(* IEC 61131-3 sources: guidance-for-physical-ai-production-designer-on-aws/source/plan2cell/crates/bt2plc/tests/golden/welding_cell_2_small/codesys/head/GVL, 2 files *)

(* ---- GVL_Cell.st ---- *)
(*
 * GVL_Cell - generated by bt2plc 0.1.0 - DO NOT EDIT
 * Plan   : bt_1790934549_welding_cell_2_small (cell welding_cell_2_small)
 * Grants : planned ticket order
 * IL01   : R1#1 W01 > R2#2 W15 > R1#3 W03 > R2#4 W10 > R1#5 W05 > R2#6 W12 > R1#7 R1_PARK > R2#7 W09
 * IL02   : R2#1 W13 > R1#2 W02 > R2#3 W14 > R1#4 W06 > R2#5 W11 > R1#6 W04 > R2#9 W07 > R1#8 HOME
 *)
{attribute 'qualified_only'}
VAR_GLOBAL CONSTANT
    (* ========================================================================
       DIMENSIONS (array bounds are literals; *_DIM >= 1)
       ======================================================================== *)
    N_ROBOTS                : INT := 2;
    N_ZONES                 : INT := 2;
    N_OPS                   : INT := 18;
    N_PREDS                 : INT := 0;

    (* ========================================================================
       PROTOCOL / TIMING
       ======================================================================== *)
    PLAN_ID                 : WORD := WORD#16#F77E;             (* fold of the plan fingerprint *)
    PROD_FOLGE              : WORD := WORD#11;                  (* default production Folge *)
    HOME_FOLGE              : WORD := WORD#125;                 (* blind homing *)
    JOB_NUMBER_BYTE         : BOOL := FALSE;                    (* FALSE: WORD LE bytes 2-3, TRUE: byte 2 *)
    PROFILE_VW              : BOOL := FALSE;                    (* TRUE: VW KS24 signal map and Folge handshake instead of the simulator telegram *)
    GRANT_POLICY            : E_GrantPolicy := E_GrantPolicy.GP_PLANNED;
    HOME_SEQUENTIAL         : BOOL := TRUE;
    AUTO_RUN                : BOOL := TRUE;                     (* start the next cycle automatically *)
    STEP_BYTE               : INT := 4;                         (* robot -> PLC, WORD LE op index *)
    REQ_BYTE                : INT := 28;                        (* robot -> PLC, DWORD LE zone requests *)
    GRANT_BYTE              : INT := 12;                        (* PLC -> robot, DWORD LE zone grants *)
    PLAN_ID_BYTE            : INT := 4;                         (* PLC -> robot, WORD LE plan id *)
    PERMIT_MASK             : DWORD := DWORD#16#80000000;       (* bit 31: permit predecessors *)
    T_RESET_PULSE           : TIME := T#1S;
    T_START_PULSE           : TIME := T#500MS;
    T_STOP_PULSE            : TIME := T#1S;
    T_HANDSHAKE             : TIME := T#5S;
    T_BRINGUP_LIMIT         : TIME := T#1M;                     (* safety enable: PROFINET connection set-up *)
    T_MISMATCH_DEBOUNCE     : TIME := T#200MS;
    T_STOP_DEBOUNCE         : TIME := T#200MS;                  (* job running: ProgRunning and ProgFinished low this long = robot stopped *)
    T_CYCLE_PAUSE           : TIME := T#2S;
    T_START_LIMIT           : TIME := T#15S;
    T_ABORT_LIMIT           : TIME := T#10S;
    T_HOME_LIMIT            : TIME := T#15S500MS;

    (* ========================================================================
       VW KS24 SIGNAL INDICES (used when PROFILE_VW; $IN/$OUT index, 1-based)
       ======================================================================== *)
    VW_READY_OUT            : INT := 9;                         (* O_R_Bereit *)
    VW_RK100_OUT            : INT := 10;                        (* O_R_RK100 safety circuit *)
    VW_AUTO_OUT             : INT := 12;                        (* O_R_Auto *)
    VW_ESTOP_OUT            : INT := 13;                        (* O_R_Notaus *)
    VW_END_OUT              : INT := 14;                        (* O_R_F_ENDE / LPKT *)
    VW_PF0_OUT              : INT := 15;                        (* O_R_PFO home position *)
    VW_STEP_OUT             : INT := 97;                        (* P_PktNr_SPS op index (16 bits) *)
    VW_REL_OUT              : INT := 41;                        (* interlock releases A41-56 *)
    VW_REQ_OUT              : INT := 81;                        (* interlock requests A81-96 *)
    VW_ERR_OUT              : INT := 225;                       (* VW_FEH_BIN_A error code (8 bits) *)
    VW_DRIVES_IN            : INT := 10;                        (* I_R_Ant_Ein *)
    VW_SRB_IN               : INT := 9;                         (* I_R_SRB Folge start *)
    VW_RESET_IN             : INT := 26;                        (* I_R_Quit_St acknowledge *)
    anInterlock             : ARRAY[1..4] OF INT := [0,0,0,0];  (* robot r, zone z -> VW interlock 1..16 (0 = not a member): index (r-1)*2+z *)

    (* ========================================================================
       ROBOTS (index = BT order)
       ======================================================================== *)
    asRobotTag              : ARRAY[1..2] OF STRING(16) := ['R1', 'R2'];
    asRobotNs               : ARRAY[1..2] OF STRING(32) := ['robot1', 'robot2'];
    abRobotActive           : ARRAY[1..2] OF BOOL := [TRUE, TRUE];
    abSafetyBypass          : ARRAY[1..2] OF BOOL := [FALSE, FALSE];(* SIMULATION ONLY: PROFIsafe slot-1 bits not required ([[robot]] safety_bypass) *)
    awRobotProdFolge        : ARRAY[1..2] OF WORD := [WORD#11, WORD#11];
    anRobotFirstOp          : ARRAY[1..2] OF INT := [1, 9];     (* op k of robot r: aOps[anRobotFirstOp[r] + k - 1] *)
    anRobotOpCount          : ARRAY[1..2] OF INT := [8, 10];

    (* ========================================================================
       ZONES - tickets of zone z: aTickets[anZoneFirst[z] .. anZoneFirst[z] + anZoneCount[z] - 1]
       ======================================================================== *)
    asZoneName              : ARRAY[1..2] OF STRING(8) := ['IL01', 'IL02'];
    anZoneFirst             : ARRAY[1..2] OF INT := [1, 9];
    anZoneCount             : ARRAY[1..2] OF INT := [8, 8];
    aTickets                : ARRAY[1..16] OF ST_Ticket := [
        (nRobot := 1, nOp := 1),    (* IL01 R1 #1 W01 *)
        (nRobot := 2, nOp := 2),    (* R2 #2 W15 *)
        (nRobot := 1, nOp := 3),    (* R1 #3 W03 *)
        (nRobot := 2, nOp := 4),    (* R2 #4 W10 *)
        (nRobot := 1, nOp := 5),    (* R1 #5 W05 *)
        (nRobot := 2, nOp := 6),    (* R2 #6 W12 *)
        (nRobot := 1, nOp := 7),    (* R1 #7 R1_PARK *)
        (nRobot := 2, nOp := 7),    (* R2 #7 W09 *)
        (nRobot := 2, nOp := 1),    (* IL02 R2 #1 W13 *)
        (nRobot := 1, nOp := 2),    (* R1 #2 W02 *)
        (nRobot := 2, nOp := 3),    (* R2 #3 W14 *)
        (nRobot := 1, nOp := 4),    (* R1 #4 W06 *)
        (nRobot := 2, nOp := 5),    (* R2 #5 W11 *)
        (nRobot := 1, nOp := 6),    (* R1 #6 W04 *)
        (nRobot := 2, nOp := 9),    (* R2 #9 W07 *)
        (nRobot := 1, nOp := 8)    (* R1 #8 HOME *)
    ];

    (* ========================================================================
       OPS - op k of robot r: aOps[anRobotFirstOp[r] + k - 1]
       ======================================================================== *)
    (* tLimit = 1.5 x tExpected + 5 s ; tZoneDeadline = 1.5 x ASAP grant + (5 + 0.2) s x depth + 10 s *)
    aOps                    : ARRAY[1..18] OF ST_OpInfo := [
        (nRobot := 1, nOp := 1, dwZoneMask := DWORD#16#00000001, nPredFirst := 0, nPredCount := 0, tExpected := T#11S132MS, tLimit := T#21S698MS, tZoneDeadline := T#10S, sName := 'W01'),    (* R1 #1 W01 *)
        (nRobot := 1, nOp := 2, dwZoneMask := DWORD#16#00000002, nPredFirst := 0, nPredCount := 0, tExpected := T#4S321MS, tLimit := T#11S482MS, tZoneDeadline := T#31S898MS, sName := 'W02'),    (* R1 #2 W02 *)
        (nRobot := 1, nOp := 3, dwZoneMask := DWORD#16#00000001, nPredFirst := 0, nPredCount := 0, tExpected := T#5S951MS, tLimit := T#13S927MS, tZoneDeadline := T#49S736MS, sName := 'W03'),    (* R1 #3 W03 *)
        (nRobot := 1, nOp := 4, dwZoneMask := DWORD#16#00000002, nPredFirst := 0, nPredCount := 0, tExpected := T#2S672MS, tLimit := T#9S8MS, tZoneDeadline := T#1M3S862MS, sName := 'W06'),    (* R1 #4 W06 *)
        (nRobot := 1, nOp := 5, dwZoneMask := DWORD#16#00000001, nPredFirst := 0, nPredCount := 0, tExpected := T#5S912MS, tLimit := T#13S868MS, tZoneDeadline := T#1M16S550MS, sName := 'W05'),    (* R1 #5 W05 *)
        (nRobot := 1, nOp := 6, dwZoneMask := DWORD#16#00000002, nPredFirst := 0, nPredCount := 0, tExpected := T#4S550MS, tLimit := T#11S825MS, tZoneDeadline := T#1M30S618MS, sName := 'W04'),    (* R1 #6 W04 *)
        (nRobot := 1, nOp := 7, dwZoneMask := DWORD#16#00000001, nPredFirst := 0, nPredCount := 0, tExpected := T#2S671MS, tLimit := T#9S7MS, tZoneDeadline := T#1M43S50MS, sName := 'R1_PARK'),    (* R1 #7 R1_PARK *)
        (nRobot := 1, nOp := 8, dwZoneMask := DWORD#16#00000002, nPredFirst := 0, nPredCount := 0, tExpected := T#8S331MS, tLimit := T#17S497MS, tZoneDeadline := T#2M25S949MS, sName := 'HOME'),    (* R1 #8 HOME *)
        (nRobot := 2, nOp := 1, dwZoneMask := DWORD#16#00000002, nPredFirst := 0, nPredCount := 0, tExpected := T#9S686MS, tLimit := T#19S529MS, tZoneDeadline := T#10S, sName := 'W13'),    (* R2 #1 W13 *)
        (nRobot := 2, nOp := 2, dwZoneMask := DWORD#16#00000001, nPredFirst := 0, nPredCount := 0, tExpected := T#8S425MS, tLimit := T#17S638MS, tZoneDeadline := T#31S898MS, sName := 'W15'),    (* R2 #2 W15 *)
        (nRobot := 2, nOp := 3, dwZoneMask := DWORD#16#00000002, nPredFirst := 0, nPredCount := 0, tExpected := T#4S724MS, tLimit := T#12S86MS, tZoneDeadline := T#49S736MS, sName := 'W14'),    (* R2 #3 W14 *)
        (nRobot := 2, nOp := 4, dwZoneMask := DWORD#16#00000001, nPredFirst := 0, nPredCount := 0, tExpected := T#4S992MS, tLimit := T#12S488MS, tZoneDeadline := T#1M3S862MS, sName := 'W10'),    (* R2 #4 W10 *)
        (nRobot := 2, nOp := 5, dwZoneMask := DWORD#16#00000002, nPredFirst := 0, nPredCount := 0, tExpected := T#5S36MS, tLimit := T#12S554MS, tZoneDeadline := T#1M16S550MS, sName := 'W11'),    (* R2 #5 W11 *)
        (nRobot := 2, nOp := 6, dwZoneMask := DWORD#16#00000001, nPredFirst := 0, nPredCount := 0, tExpected := T#4S821MS, tLimit := T#12S232MS, tZoneDeadline := T#1M30S618MS, sName := 'W12'),    (* R2 #6 W12 *)
        (nRobot := 2, nOp := 7, dwZoneMask := DWORD#16#00000001, nPredFirst := 0, nPredCount := 0, tExpected := T#2S699MS, tLimit := T#9S48MS, tZoneDeadline := T#1M52S256MS, sName := 'W09'),    (* R2 #7 W09 *)
        (nRobot := 2, nOp := 8, dwZoneMask := DWORD#16#00000000, nPredFirst := 0, nPredCount := 0, tExpected := T#4S594MS, tLimit := T#11S891MS, tZoneDeadline := T#2M1S505MS, sName := 'W08'),    (* R2 #8 W08 *)
        (nRobot := 2, nOp := 9, dwZoneMask := DWORD#16#00000002, nPredFirst := 0, nPredCount := 0, tExpected := T#4S769MS, tLimit := T#12S154MS, tZoneDeadline := T#2M13S596MS, sName := 'W07'),    (* R2 #9 W07 *)
        (nRobot := 2, nOp := 10, dwZoneMask := DWORD#16#00000000, nPredFirst := 0, nPredCount := 0, tExpected := T#6S229MS, tLimit := T#14S344MS, tZoneDeadline := T#2M25S949MS, sName := 'HOME')    (* R2 #10 HOME *)
    ];

    (* ========================================================================
       PERMIT PREDECESSORS - op preds: aPreds[nPredFirst .. nPredFirst + nPredCount - 1]
       ======================================================================== *)
    aPreds                  : ARRAY[1..1] OF ST_Ticket := [
        (nRobot := 0, nOp := 0)    (* no permit predecessors *)
    ];
END_VAR

(* ---- GVL_IO.st ---- *)
(*
 * GVL_IO - Head PLC I/O, one block per robot
 * Generated by bt2plc 0.1.0 for cell welding_cell_2_small (plan bt_1790934549_welding_cell_2_small)
 *
 * This is the PROFINET Controller (master) side.
 * From the controller's perspective:
 *   "Inputs"  = data received FROM the robot device (robot status)
 *   "Outputs" = data sent TO the robot device (PLC commands)
 *
 * Map in the I/O Mapping tab of each KUKA device under the PN-Controller:
 *   SafeIO_FDIO64_<tag> inputs  -> bySafeIn0_<tag>..bySafeIn7_<tag>
 *   SafeIO_FDIO64_<tag> outputs -> bySafeOut0_<tag>..bySafeOut7_<tag>
 *   VASS_DIO256_<tag> inputs    -> aVassInputData_<tag>
 *   VASS_DIO256_<tag> outputs   -> aVassOutputData_<tag>
 *
 * Only PLC_PRG accesses this GVL: whole arrays and single bytes are copied
 * into / out of FB_Cell (never write single elements of these arrays).
 *)

{attribute 'qualified_only'}
VAR_GLOBAL

    (* ========================================================================
       R1 - robot1 - kuka_robi1 (kuka-robi1, 192.168.100.11)
       ======================================================================== *)

    (* SLOT 1 - PROFIsafe FDIO64: safe status FROM robot (8 bytes) *)
    bySafeIn0_R1            : BYTE;     (* Byte 0: Drives OK, Stopped, Reduced speed... *)
    bySafeIn1_R1            : BYTE;     (* Byte 1: Gates, E-Stop, Enabling... *)
    bySafeIn2_R1            : BYTE;     (* Byte 2: STO, SS1, SS2, SOS, SLS... *)
    bySafeIn3_R1            : BYTE;
    bySafeIn4_R1            : BYTE;
    bySafeIn5_R1            : BYTE;
    bySafeIn6_R1            : BYTE;
    bySafeIn7_R1            : BYTE;

    (* SLOT 1 - PROFIsafe FDIO64: safe commands TO robot (8 bytes) *)
    bySafeOut0_R1           : BYTE;     (* Byte 0: Drive enable, E-Stop, SS1, SS2, SLS... *)
    bySafeOut1_R1           : BYTE;     (* Byte 1: Zone enables *)
    bySafeOut2_R1           : BYTE;
    bySafeOut3_R1           : BYTE;
    bySafeOut4_R1           : BYTE;
    bySafeOut5_R1           : BYTE;
    bySafeOut6_R1           : BYTE;
    bySafeOut7_R1           : BYTE;

    (* SLOT 2 - DIO256 VASS telegram (32 bytes each direction) *)
    aVassInputData_R1       : ARRAY[0..31] OF BYTE;         (* VASS status FROM robot *)
    aVassOutputData_R1      : ARRAY[0..31] OF BYTE;         (* VASS commands TO robot *)

    (* ========================================================================
       R2 - robot2 - kuka_robi2 (kuka-robi2, 192.168.100.12)
       ======================================================================== *)

    (* SLOT 1 - PROFIsafe FDIO64: safe status FROM robot (8 bytes) *)
    bySafeIn0_R2            : BYTE;     (* Byte 0: Drives OK, Stopped, Reduced speed... *)
    bySafeIn1_R2            : BYTE;     (* Byte 1: Gates, E-Stop, Enabling... *)
    bySafeIn2_R2            : BYTE;     (* Byte 2: STO, SS1, SS2, SOS, SLS... *)
    bySafeIn3_R2            : BYTE;
    bySafeIn4_R2            : BYTE;
    bySafeIn5_R2            : BYTE;
    bySafeIn6_R2            : BYTE;
    bySafeIn7_R2            : BYTE;

    (* SLOT 1 - PROFIsafe FDIO64: safe commands TO robot (8 bytes) *)
    bySafeOut0_R2           : BYTE;     (* Byte 0: Drive enable, E-Stop, SS1, SS2, SLS... *)
    bySafeOut1_R2           : BYTE;     (* Byte 1: Zone enables *)
    bySafeOut2_R2           : BYTE;
    bySafeOut3_R2           : BYTE;
    bySafeOut4_R2           : BYTE;
    bySafeOut5_R2           : BYTE;
    bySafeOut6_R2           : BYTE;
    bySafeOut7_R2           : BYTE;

    (* SLOT 2 - DIO256 VASS telegram (32 bytes each direction) *)
    aVassInputData_R2       : ARRAY[0..31] OF BYTE;         (* VASS status FROM robot *)
    aVassOutputData_R2      : ARRAY[0..31] OF BYTE;         (* VASS commands TO robot *)

END_VAR
